// TwinCAT 3 PLC project Storage_Main
// ProgramVersion: 3.1.4026.27
// libraries:
//   CmpBitmapPool, * (System)
//   Tc2_Standard, * (Beckhoff Automation GmbH)
//   Tc2_System, * (Beckhoff Automation GmbH)
//   Tc3_Module, * (Beckhoff Automation GmbH)
//   VisuSymbols,3.5.10.0,System
// project tree:
//   / GlobalTextList.TcGTLO, PlcTask.TcTTO, Visualization Manager.TcVMO (not stored), VISU_TASK.TcTTO
//   POUs/ MAIN.TcPOU
//   VISUs/ Billeder.TcIPO (not stored), IO.TcVIS, Start.TcVIS
// real-time tasks:
//   TASK PlcTask: cycle T#10ms, priority 20, ADS port 350
//   TASK VISU_TASK: cycle T#200000us, priority 30, ADS port 351
// motion (NC):
//   TASK EncoderHorizontal SAF: cycle T#2ms, priority 4, ADS port 501
//   TASK EncoderHorizontal SVB: cycle T#10ms, priority 8, ADS port 511
//   AXIS X (id 1)
//     OtherSettings: AllowMotionCmdToSlave=true
//     encoder EncType=1
//     drive DrvType=5
//       Analog: TorqueSetpointScale=10, ScaleFactorActTorque=0.1
//     controller CtrType=1
//       CtrPara: PriorControlFactor=1
//         Observer: BandWidth=20
// I/O:
//   DEVICE Device 1 (EtherCAT Automation Protocol), AmsNetId 10.180.10.242.2.1
//   DEVICE Device 3 (EtherCAT), AmsNetId 10.180.10.242.4.1
//     Term 1 (EK1100) [EK1100 EtherCAT Coupler (2A E-Bus)]
//       Term 2 (EL1202) [EL1202 2Ch. Fast Dig. Input 24V, 1µs]
//       Term 3 (EL1202) [EL1202 2Ch. Fast Dig. Input 24V, 1µs]
//       Term 4 (EL1008) [EL1008 8Ch. Dig. Input 24V, 3ms]
//       Term 5 (EL1008) [EL1008 8Ch. Dig. Input 24V, 3ms]
//       Term 6 (EL2008) [EL2008 8Ch. Dig. Output 24V, 0.5A]
//       Term 7 (EL3064) [EL3064 4Ch. Ana. Input 0-10V]
//       Term 8 (EL4022) [EL4022 2Ch. Ana. Output 4-20mA, 12bit]
//       Term 9 (EL3072) [EL3072 2Ch. Ana. Input +/-10V, +/-20mA]
//       Term 10 (EL6631-0010) [EL6631-0010 PROFINET IO Device]
//       Term 11 (EL9011) [EL9011 End Terminal]
// variable links:
//   Storage_Main/Storage_Main Instance <-> Device 3 (EtherCAT)/Term 1 (EK1100)/Term 2 (EL1202)
//     PlcTask Inputs/MAIN.B5 <-> Channel 1/MAIN.B5
//     PlcTask Inputs/MAIN.B6 <-> Channel 2/MAIN.B6
//   Storage_Main/Storage_Main Instance <-> Device 3 (EtherCAT)/Term 1 (EK1100)/Term 3 (EL1202)
//     PlcTask Inputs/MAIN.B3 <-> Channel 1/MAIN.B3
//     PlcTask Inputs/MAIN.B4 <-> Channel 2/MAIN.B4
//   Storage_Main/Storage_Main Instance <-> Device 3 (EtherCAT)/Term 1 (EK1100)/Term 4 (EL1008)
//     PlcTask Inputs/MAIN.B1 <-> Channel 1/MAIN.B1
//     PlcTask Inputs/MAIN.B2 <-> Channel 2/MAIN.B2
//     PlcTask Inputs/MAIN.B7 <-> Channel 3/Input
//     PlcTask Inputs/MAIN.B8 <-> Channel 4/Input
//   Storage_Main/Storage_Main Instance <-> Device 3 (EtherCAT)/Term 1 (EK1100)/Term 5 (EL1008)
//     PlcTask Inputs/MAIN.B10 <-> Channel 2/Input
//     PlcTask Inputs/MAIN.B9 <-> Channel 1/Input
//   Storage_Main/Storage_Main Instance <-> Device 3 (EtherCAT)/Term 1 (EK1100)/Term 6 (EL2008)
//     PlcTask Outputs/MAIN.M1_Back <-> Channel 2/Output
//     PlcTask Outputs/MAIN.M2_Back <-> Channel 4/Output
//     PlcTask Outputs/MAIN.M4_Back <-> Channel 8/Output
//     PlcTask Outputs/MAIN.M1_Forward <-> Channel 1/Output
//     PlcTask Outputs/MAIN.M2_Forward <-> Channel 3/Output
//     PlcTask Outputs/MAIN.M4_Forward <-> Channel 7/Output
//     PlcTask Outputs/MAIN.M3_Down <-> Channel 5/Output
//     PlcTask Outputs/MAIN.M3_Up <-> Channel 6/Output

CONFIGURATION Storage_Main
    RESOURCE PLC ON TwinCAT3
        TASK PlcTask(INTERVAL := T#10ms, PRIORITY := 20);
        TASK VISU_TASK(INTERVAL := T#200000us, PRIORITY := 30);
        PROGRAM MAIN WITH PlcTask : MAIN;
        PROGRAM VisuElems_Visu_Prg WITH VISU_TASK : VisuElems.Visu_Prg;
    END_RESOURCE
END_CONFIGURATION

// ---- POUs/MAIN.TcPOU
PROGRAM MAIN
VAR
    // ---------------- INPUTS ----------------
    B1  AT %I* : BOOL;  // Nr. 5,  B1: reference switch horizontal axis
    B2  AT %I* : BOOL;  // Nr. 6,  B2: light-barrier inside
    B3  AT %I* : BOOL;  // Nr. 7,  B3: light-barrier outside
    B4  AT %I* : BOOL;  // Nr. 8,  B4: reference switch vertical axis
    B5  AT %I* : BOOL;  // Nr. 11, B5: encoder horizontal axis impulse 1  (EL1202 ch. 1)
    B6  AT %I* : BOOL;  // Nr. 12, B6: encoder horizontal axis impulse 2  (EL1202 ch. 2)
    B7  AT %I* : BOOL;  // Nr. 13, B7: encoder vertical axis impulse 1
    B8  AT %I* : BOOL;  // Nr. 14, B8: encoder vertical axis impulse 2
    B9  AT %I* : BOOL;  // Nr. 15, B9: reference switch cantilever front
    B10 AT %I* : BOOL;  // Nr. 16, B10: reference switch cantilever back

    // Optional push buttons (not in the I/O list - leave unlinked if not used)
    bButtonHoming AT %I* : BOOL;  // Start homing
    bButtonMove   AT %I* : BOOL;  // Move to xPosition[nSlot]
    bButtonStop   AT %I* : BOOL;  // Stop (level: stops as long as pressed)

    // ---------------- OUTPUTS ----------------
    M1_Forward AT %Q* : BOOL;  // Nr. 17, Q1 (M1): motor conveyor belt forward
    M1_Back    AT %Q* : BOOL;  // Nr. 18, Q2 (M1): motor conveyor belt backward
    M2_Forward AT %Q* : BOOL;  // Nr. 19, Q3 (M2): motor horizontal towards rack
    M2_Back    AT %Q* : BOOL;  // Nr. 20, Q4 (M2): motor horizontal towards conveyor belt
    M3_Down    AT %Q* : BOOL;  // Nr. 21, Q5 (M3): motor vertical axis downward
    M3_Up      AT %Q* : BOOL;  // Nr. 22, Q6 (M3): motor vertical axis upward
    M4_Forward AT %Q* : BOOL;  // Nr. 23, Q7 (M4): motor cantilever forward
    M4_Back    AT %Q* : BOOL;  // Nr. 24, Q8 (M4): motor cantilever backward

    // ---------------- POSITIONS (horizontal / X axis) ----------------
    // Rack columns in encoder counts: [1] = column 1, [2] = column 2, [3] = column 3
    xPosition : ARRAY[1..3] OF DINT := [185, 365, 545];
    nSlot     : INT := 1;       // Which column to move to / teach (1..3)
    bTeach    : BOOL;           // Save current nPosition into xPosition[nSlot]

    // ---------------- COMMANDS (horizontal / X axis) ----------------
    // Set online with "Write values" / Ctrl+F7
    bJogForward  : BOOL;            // Manual move towards rack (step 0 only)
    bJogBackward : BOOL;            // Manual move towards conveyor (step 0 only)
    bStartHoming : BOOL;            // Start homing sequence
    bStartMove   : BOOL;            // Move to xPosition[nSlot]
    bStop        : BOOL;            // Stop everything
    nTarget      : DINT;            // Current target (set from xPosition)
    nTolerance   : DINT := 5;       // Deadband in counts

    // ---------------- EDGE DETECTION ----------------
    rtHoming : R_TRIG;
    rtMove   : R_TRIG;

    // ---------------- ENCODER (horizontal / X axis) ----------------
    nState      : BYTE;             // Current state 0..3
    nPrevState  : BYTE;             // State in previous cycle
    bInit       : BOOL := TRUE;     // First cycle flag
    nPosition   : DINT;             // Position in counts (300 per output shaft rev.)
    nErrorCount : UDINT;            // Number of missed states

    // ---------------- SEQUENCE / STATUS ----------------
    nStep       : INT := 0;         // 0 = idle, 10 = homing, 20 = moving to target
    bHomed      : BOOL;             // TRUE when zero point is found
    bInPosition : BOOL;             // TRUE when target is reached
	// counter
	totalValue: INT;
	
	counterB1  : DINT;
	counterB2  : DINT;
	counterB3  : DINT;
	counterB4  : DINT;
	counterB5  : DINT;
	counterB6  : DINT;
	counterB7  : DINT;
	counterB8  : DINT;
	counterB9  : DINT;
	counterB10 : DINT;
END_VAR

Test();

ACTION Test:
// =====================================================
// 1. ENCODER: count up/down based on B5 (A) and B6 (B)
// =====================================================
nState := 0;                                        // default: A=0, B=0
IF B5 AND NOT B6 THEN nState := 1; END_IF           // A=1, B=0
IF B5 AND B6 THEN nState := 2; END_IF               // A=1, B=1
IF NOT B5 AND B6 THEN nState := 3; END_IF           // A=0, B=1

IF B1 THEN
    counterB1 := counterB1 + 1;
END_IF
IF B2 THEN
    counterB2 := counterB2 + 1;
END_IF
IF B3 THEN
    counterB3 := counterB3 + 1;
END_IF
IF B4 THEN
    counterB4 := counterB4 + 1;
END_IF
IF B5 THEN
    counterB5 := counterB5 + 1;
END_IF
IF B6 THEN
    counterB6 := counterB6 + 1;
END_IF
IF B7 THEN
    counterB7 := counterB7 + 1;
END_IF
IF B8 THEN
    counterB8 := counterB8 + 1;
END_IF
IF B9 THEN
    counterB9 := counterB9 + 1;
END_IF
IF B10 THEN
    counterB10 := counterB10 + 1;
END_IF

CASE (nState + 4 - nPrevState) MOD 4 OF
    1: nPosition := nPosition + 1;                  // one step forward
    3: nPosition := nPosition - 1;                  // one step backward
    2: nErrorCount := nErrorCount + 1;              // state missed
END_CASE

nPrevState := nState;


// =====================================================
// 2. PUSH BUTTONS: edge detection -> commands
// =====================================================
rtHoming(CLK := bButtonHoming);
rtMove(CLK := bButtonMove);

IF rtHoming.Q THEN bStartHoming := TRUE; END_IF     // TRUE for one cycle only
IF rtMove.Q THEN bStartMove := TRUE; END_IF
IF bButtonStop THEN bStop := TRUE; END_IF           // level: no edge needed


// =====================================================
// 3. STOP: always returns to step 0
// =====================================================
IF bStop THEN
    bStop := FALSE;
    bStartHoming := FALSE;
    bStartMove := FALSE;
    nStep := 0;
END_IF


// =====================================================
// 4. TEACH: save current position into the array
// =====================================================
IF bTeach THEN
    bTeach := FALSE;
    IF bHomed AND nSlot >= 1 AND nSlot <= 3 THEN
        xPosition[nSlot] := nPosition;
    END_IF
END_IF


// =====================================================
// 5. SEQUENCE (horizontal / X axis, motor M2)
// =====================================================
CASE nStep OF

    0:  // ----- Idle: manual jog only -----
        M2_Forward := bJogForward AND NOT bJogBackward;
        M2_Back    := bJogBackward AND NOT bJogForward AND NOT B1;

        IF bStartHoming THEN
            bStartHoming := FALSE;
            bHomed := FALSE;
            nStep := 10;
        END_IF

        IF bStartMove THEN
            bStartMove := FALSE;
            IF bHomed AND nSlot >= 1 AND nSlot <= 3 THEN
                nTarget := xPosition[nSlot];        // look up target in the array
                bInPosition := FALSE;
                nStep := 20;
            END_IF
        END_IF

    10: // ----- Homing: move towards conveyor until reference switch B1 -----
        M2_Forward := FALSE;
        M2_Back    := TRUE;

        IF B1 THEN                                  // level, not edge
            M2_Back := FALSE;
            nPosition := 0;                         // zero point = where the switch triggers
            bHomed := TRUE;
            nStep := 0;
        END_IF

    20: // ----- Move to nTarget -----
        M2_Forward := FALSE;                        // default: motor off
        M2_Back    := FALSE;

        IF nPosition < nTarget - nTolerance THEN
            M2_Forward := TRUE;                     // too close to conveyor -> towards rack
        END_IF

        IF nPosition > nTarget + nTolerance THEN
            M2_Back := TRUE;                        // too far towards rack -> towards conveyor
        END_IF

        IF NOT M2_Forward AND NOT M2_Back THEN
            bInPosition := TRUE;                    // within tolerance -> done
            nStep := 0;
        END_IF

END_CASE


// =====================================================
// 6. SAFETY: never both directions at the same time
// =====================================================
IF M2_Forward AND M2_Back THEN
    M2_Forward := FALSE;
    M2_Back    := FALSE;
END_IF
END_ACTION

END_PROGRAM

// ---- GlobalTextList.TcGTLO
TEXTLIST GlobalTextList
  737 = 'Arm Back'
  219 = 'Arm Down'
  893 = 'Arm Forward'
  973 = 'B1'
  905 = 'B10'
  806 = 'B2'
  287 = 'B3'
  334 = 'B4'
  502 = 'B5'
  579 = 'B6'
  213 = 'B7'
  974 = 'B8'
  734 = 'B9'
  283 = 'Back'
  163 = 'Crane Back'
  196 = 'Crane Down'
  176 = 'Crane Forward'
  61 = 'Crane Up'
  422 = 'Emne Frem'
  568 = 'Emne Tilbage'
  629 = 'Feed the packman'
  939 = 'Feed the Pacman'
  826 = 'Forward'
  910 = 'Settings'
  77 = 'Slay the demon'
  19 = 'Start'
  1 = 'TEST'
END_TEXTLIST

// ---- VISUs/IO.TcVIS
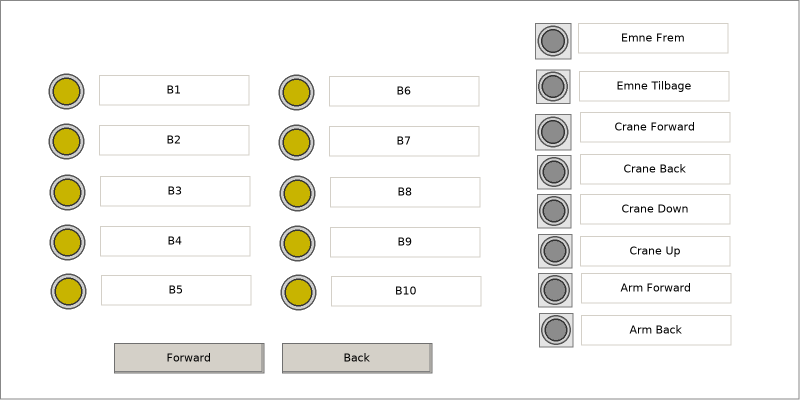
VISUALIZATION IO  // 800x400
    Lamp1 (46,71 41x41), variable: MAIN.B1, style: Lamp-Lamp1-Yellow
    Textfield (99,75 150x30), "B1"
    Textfield (99,125 150x30), "B2"
    Lamp1 (46,121 41x41), variable: MAIN.B2, style: Lamp-Lamp1-Yellow
    Lamp1 (47,172 41x41), variable: MAIN.B3, style: Lamp-Lamp1-Yellow
    Textfield (100,176 150x30), "B3"
    Textfield (100,226 150x30), "B4"
    Lamp1 (47,222 41x41), variable: MAIN.B4, style: Lamp-Lamp1-Yellow
    Lamp1 (48,271 41x41), variable: MAIN.B5, style: Lamp-Lamp1-Yellow
    Textfield (101,275 150x30), "B5"
    Lamp1 (276,72 41x41), variable: MAIN.B6, style: Lamp-Lamp1-Yellow
    Textfield (329,76 150x30), "B6"
    Textfield (329,126 150x30), "B7"
    Lamp1 (276,122 41x41), variable: MAIN.B7, style: Lamp-Lamp1-Yellow
    Lamp1 (277,173 41x41), variable: MAIN.B8, style: Lamp-Lamp1-Yellow
    Textfield (330,177 150x30), "B8"
    Textfield (330,227 150x30), "B9"
    Lamp1 (277,223 41x41), variable: MAIN.B9, style: Lamp-Lamp1-Yellow
    Lamp1 (278,272 41x41), variable: MAIN.B10, style: Lamp-Lamp1-Yellow
    Textfield (331,276 150x30), "B10"
    Textfield (579,71 150x30), "Emne Tilbage"
    PushSwitch (536,69 34x35), variable: MAIN.M1_Forward, behaviour: TAP, style: Switch-PushSwitch-Gray
    PushSwitch (535,23 36x36), variable: MAIN.M1_Back, behaviour: TAP, style: Switch-PushSwitch-Gray
    Textfield (578,23 150x30), "Emne Frem"
    Textfield (580,112 150x30), "Crane Forward"
    PushSwitch (535,114 36x36), variable: MAIN.M2_Forward, behaviour: TAP, style: Switch-PushSwitch-Gray
    PushSwitch (537,155 34x34), variable: MAIN.M2_Back, behaviour: TAP, style: Switch-PushSwitch-Gray
    Textfield (580,154 150x30), "Crane Back"
    Textfield (580,194 150x30), "Crane Down"
    PushSwitch (537,194 34x34), variable: MAIN.M3_Down, behaviour: TAP, style: Switch-PushSwitch-Gray
    PushSwitch (538,234 34x34), variable: MAIN.M3_Up, behaviour: TAP, style: Switch-PushSwitch-Gray
    Textfield (580,236 150x30), "Crane Up"
    Textfield (581,273 150x30), "Arm Forward"
    PushSwitch (538,273 34x34), variable: MAIN.M4_Forward, behaviour: TAP, style: Switch-PushSwitch-Gray
    PushSwitch (539,313 34x34), variable: MAIN.M4_Back, behaviour: TAP, style: Switch-PushSwitch-Gray
    Textfield (581,315 150x30), "Arm Back"
    Button (114,343 150x30), "Forward"
        tap MAIN.bJogForward
    Button (282,343 150x30), "Back"
        tap MAIN.bJogBackward
END_VISUALIZATION

// ---- VISUs/Start.TcVIS
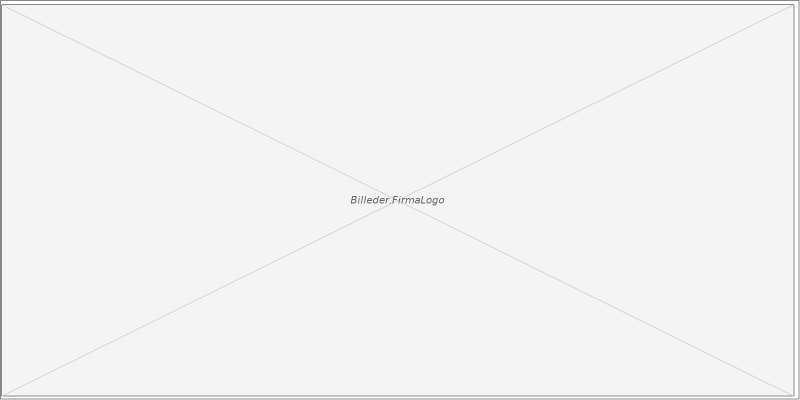
VISUALIZATION Start  // 800x400
    Image (1,4 793x392), image: Billeder.FirmaLogo
END_VISUALIZATION
